(* IEC 61131-3 sources: plcassist-cli/packages/volt-lsp-iec/test-corpus/pro2193/Device/Plc Logic/Application/09 Misc/Library Manager/CmpSchedule, 15 files *)

(* ---- SCHEDGETCURRENTTASK.fun ---- *)
FUNCTION SCHEDGETCURRENTTASK : RTS_IEC_HANDLE
VAR_INPUT
	PRESULT : POINTER TO RTS_IEC_RESULT;
END_VAR
END_FUNCTION

(* ---- SCHEDGETNUMOFTASKS.fun ---- *)
FUNCTION SCHEDGETNUMOFTASKS : DINT
VAR_INPUT
	PAPP : POINTER TO APPLICATION;
	PRESULT : POINTER TO RTS_IEC_RESULT;
END_VAR
END_FUNCTION

(* ---- SCHEDGETPROCESSORLOAD.fun ---- *)
FUNCTION SCHEDGETPROCESSORLOAD : UDINT
VAR_INPUT
	PRESULT : POINTER TO RTS_IEC_RESULT;
END_VAR
END_FUNCTION

(* ---- SCHEDGETTASKEVENTBYHANDLE.fun ---- *)
FUNCTION SCHEDGETTASKEVENTBYHANDLE : RTS_IEC_HANDLE
VAR_INPUT
	HSCHEDTASK : RTS_IEC_HANDLE;
	PRESULT : POINTER TO RTS_IEC_RESULT;
END_VAR
END_FUNCTION

(* ---- SCHEDGETTASKHANDLEBYINDEX.fun ---- *)
FUNCTION SCHEDGETTASKHANDLEBYINDEX : RTS_IEC_HANDLE
VAR_INPUT
	PAPP : POINTER TO APPLICATION;
	NINDEX : DINT;
	PRESULT : POINTER TO RTS_IEC_RESULT;
END_VAR
END_FUNCTION

(* ---- SCHEDGETTASKHANDLEBYNAME.fun ---- *)
FUNCTION SCHEDGETTASKHANDLEBYNAME : RTS_IEC_HANDLE
VAR_INPUT
	PRESULT : POINTER TO RTS_IEC_RESULT;
END_VAR
VAR_IN_OUT
	PSZTASKNAME : STRING;
END_VAR
END_FUNCTION

(* ---- SCHEDGETTASKINTERVAL.fun ---- *)
FUNCTION SCHEDGETTASKINTERVAL : RTS_IEC_RESULT
VAR_INPUT
	HSCHEDTASK : RTS_IEC_HANDLE;
END_VAR
VAR_IN_OUT
	PULINTERVAL : UDINT;
END_VAR
END_FUNCTION

(* ---- SCHEDPOSTEXTERNALEVENT.fun ---- *)
FUNCTION SCHEDPOSTEXTERNALEVENT : RTS_IEC_RESULT
VAR_INPUT
	HEXTEVENT : RTS_IEC_HANDLE;
END_VAR
END_FUNCTION

(* ---- SCHEDREGISTEREXTERNALEVENT.fun ---- *)
FUNCTION SCHEDREGISTEREXTERNALEVENT : RTS_IEC_HANDLE
VAR_INPUT
	PSZEXTEVENTNAME : REFERENCE TO STRING;
	PRESULT : POINTER TO RTS_IEC_RESULT;
END_VAR
END_FUNCTION

(* ---- SCHEDSETTASKINTERVAL.fun ---- *)
FUNCTION SCHEDSETTASKINTERVAL : RTS_IEC_RESULT
VAR_INPUT
	HSCHEDTASK : RTS_IEC_HANDLE;
	ULINTERVAL : UDINT;
END_VAR
END_FUNCTION

(* ---- SCHEDTASKRESUME.fun ---- *)
FUNCTION SCHEDTASKRESUME : SysTypes.RTS_IEC_RESULT
VAR_INPUT
	HSCHEDTASK : SysTypes.RTS_IEC_HANDLE;
END_VAR
END_FUNCTION

(* ---- SCHEDTASKSUSPEND.fun ---- *)
FUNCTION SCHEDTASKSUSPEND : SysTypes.RTS_IEC_RESULT
VAR_INPUT
	HSCHEDTASK : SysTypes.RTS_IEC_HANDLE;
END_VAR
END_FUNCTION

(* ---- SCHEDUNREGISTEREXTERNALEVENT.fun ---- *)
FUNCTION SCHEDUNREGISTEREXTERNALEVENT : RTS_IEC_RESULT
VAR_INPUT
	HEXTEVENT : RTS_IEC_HANDLE;
END_VAR
END_FUNCTION

(* ---- SCHEDWAITBUSY.fun ---- *)
FUNCTION SCHEDWAITBUSY : RTS_IEC_RESULT
VAR_IN_OUT
	PTSLEEPUS : SYSTIME;
END_VAR
END_FUNCTION

(* ---- SCHEDWAITSLEEP.fun ---- *)
FUNCTION SCHEDWAITSLEEP : RTS_IEC_RESULT
VAR_IN_OUT
	PTSLEEPUS : SYSTIME;
END_VAR
END_FUNCTION
